FUNCTION_BLOCK AQ_BYTE_TO_Q (* Composite FB for convert BYTE (QUARTER, 2 Bit) to AQ *)
  (* Standard: 61499-2; Description: Copyright (c) 2026 HR Agrartechnik GmbH This program and the accompanying materials are made available under the terms of the Eclipse Public License 2.0 which is available at https://www.eclipse.org/legal/epl-2.0/ SPDX-License-Identifier: EPL-2.0 *)
  (* Version 1.0, 2026-11-13, Franz Höpfinger, HR Agrartechnik GmbH, Initial Version - Luecke geschlossen (analog zu AB_BYTE_TO_B) *)
  PACKAGE adapter::conversion::unidirectional;
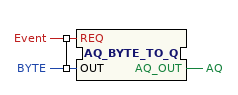
  EVENT_INPUT
    REQ WITH OUT; (* Request to Adapter *)
  END_EVENT
  VAR_INPUT
    OUT : BYTE; (* Output data to Adapter *)
  END_VAR
  PLUGS
    AQ_OUT : adapter::types::unidirectional::AQ; (* Adapter Output *)
  END_PLUGS
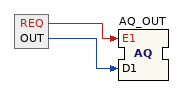
  EVENT_CONNECTIONS
    REQ TO AQ_OUT.E1;
  END_CONNECTIONS
  DATA_CONNECTIONS
    OUT TO AQ_OUT.D1;
  END_CONNECTIONS
END_FUNCTION_BLOCK
